Fanuc KAREL source: KB00149.KL

PROGRAM KB00149
%NOLOCKGROUP
%ENVIRONMENT MOTN
VAR
  P1: BOOLEAN
BEGIN
  P1 = TRUE
  RESET(P1)
END KB00149
